SUBAPPLICATION Uebung_094b3e_AX (* Wie Uebung_094b3_AX, aber mit dritter Gruppe OptionalGroup_001b, die ueber AOption_T_2 (Abgriff hinter 001 und 002) und AOption_OR_2 aktiv ist, sobald 001 ODER 002 aktiv ist (K=2 oder K=3) - bei K=1 (DummyGroup) bleibt sie aus. *)
  (* Standard: 61499-2; Description: Copyright (c) 2026 Meisterschulen am Ostbahnhof This program and the accompanying materials are made available under the terms of the Eclipse Public License 2.0 which is available at https://www.eclipse.org/legal/epl-2.0/ SPDX-License-Identifier: EPL-2.0 *)
  (* Version 1.0, 2026-10-17, Franz Höpfinger, Meisterschulen am Ostbahnhof, Kopie von Uebung_094b3_AX mit dritter Gruppe (001b) hinter 001 und 002 per T-Stueck + OR, nicht bei DummyGroup. *)
  PACKAGE Uebungen;
  IMPORT Uebungen::const::UT::DefaultPool::InputNumber_I1;
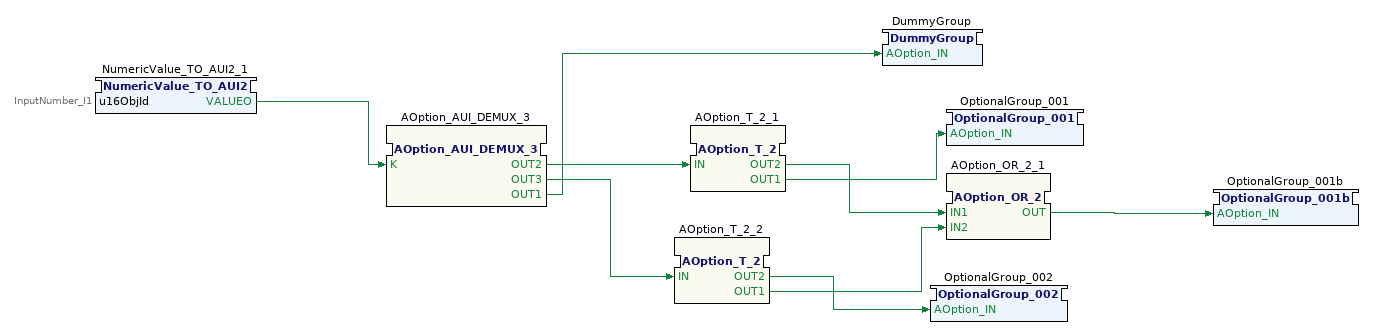
  FBS
    AOption_AUI_DEMUX_3 : Option::selection::AOption_AUI_DEMUX_3;
    AOption_T_2_1 : Option::splitting::AOption_T_2;
    AOption_T_2_2 : Option::splitting::AOption_T_2;
    AOption_OR_2_1 : Option::merging::AOption_OR_2;
  END_FBS
  SUBAPPS
    NumericValue_TO_AUI2_1 : MyLib::sys::NumericValue_TO_AUI2(u16ObjId := InputNumber_I1);
    OptionalGroup_001 : MyLib_AX_Option::sys::OptionalGroup_001;
    OptionalGroup_002 : MyLib_AX_Option::sys::OptionalGroup_002;
    OptionalGroup_001b : MyLib_AX_Option::sys::OptionalGroup_001b;
    DummyGroup : MyLib_AX_Option::sys::DummyGroup;
  END_SUBAPPS
  ADAPTER_CONNECTIONS
    NumericValue_TO_AUI2_1.VALUEO TO AOption_AUI_DEMUX_3.K;
    AOption_AUI_DEMUX_3.OUT2 TO AOption_T_2_1.IN;
    AOption_T_2_1.OUT2 TO AOption_OR_2_1.IN1;
    AOption_AUI_DEMUX_3.OUT3 TO AOption_T_2_2.IN;
    AOption_T_2_2.OUT2 TO OptionalGroup_002.AOption_IN;
    AOption_T_2_2.OUT1 TO AOption_OR_2_1.IN2;
    AOption_OR_2_1.OUT TO OptionalGroup_001b.AOption_IN;
    AOption_AUI_DEMUX_3.OUT1 TO DummyGroup.AOption_IN;
    AOption_T_2_1.OUT1 TO OptionalGroup_001.AOption_IN;
  END_CONNECTIONS
END_SUBAPPLICATION
